// TIA Portal V21 export
// export: Created 2026-08-21T20:18:51.0501839Z, ExportSetting None, DisplayName Totally Integrated Automation Portal, DisplayVersion V21, DisplayName STEP 7 Professional, DisplayVersion V21, DisplayName STEP 7 Safety, DisplayVersion V21, DisplayName Tech WebApplication, DisplayVersion V21, DisplayName WinCC Basic/Comfort/Advanced, DisplayVersion V21, DisplayName WinCC Professional, DisplayVersion V21, DisplayName WinCC Unified, DisplayVersion V21
FUNCTION "V100" : Void   // FC3, FBD
{ S7_Optimized_Access := 'TRUE' }
// stored: SetENOAutomatically false
   VAR_TEMP
      Temp : "DigVal";
      In03 : "DigVal";
      Temp_FF : "DigVal";
      Temp_fromCTRL : "StruCm";
   END_VAR
BEGIN

REGION Network 1: VlvAnL interconnections
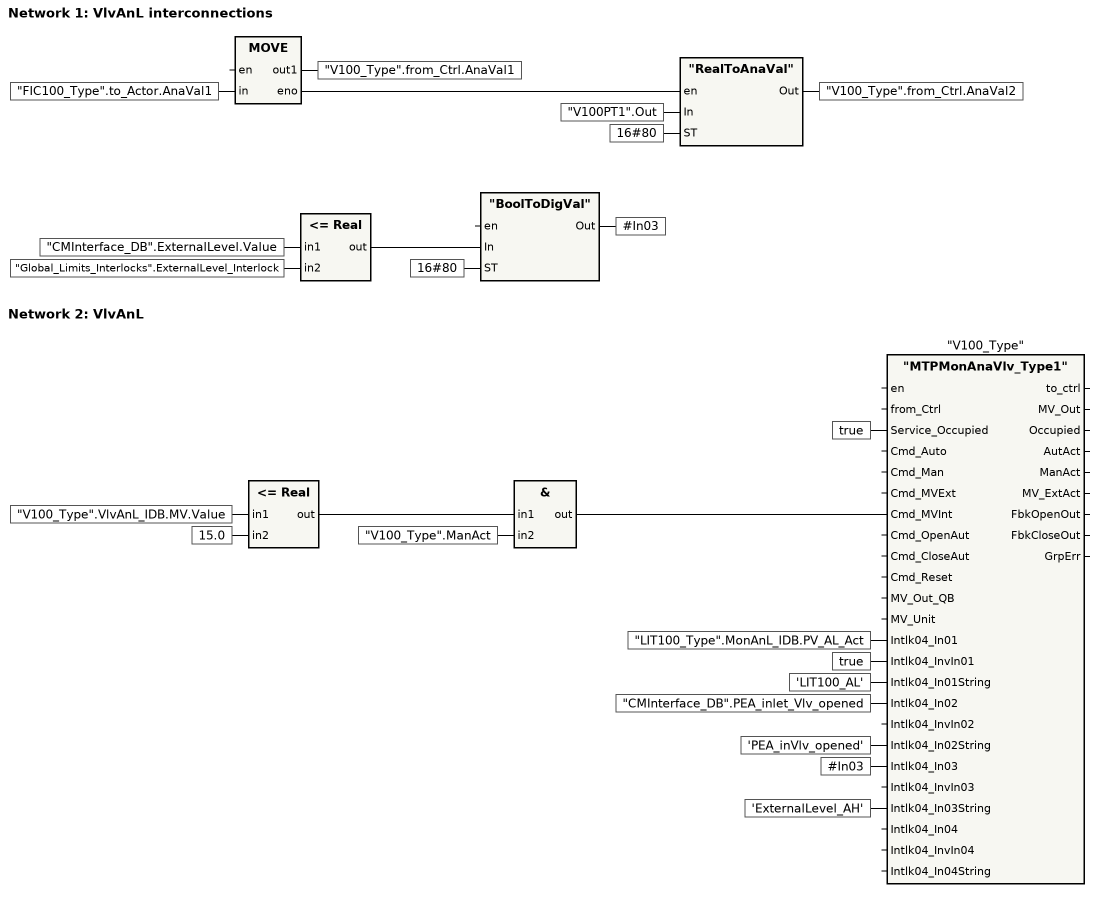
   "V100_Type".from_Ctrl.AnaVal1 := "FIC100_Type".to_Actor.AnaVal1;
   "RealToAnaVal"(In := "V100PT1".Out, ST := 16#80, Out => "V100_Type".from_Ctrl.AnaVal2);
   "BoolToDigVal"(In := "CMInterface_DB".ExternalLevel.Value <= "Global_Limits_Interlocks".ExternalLevel_Interlock,
                  ST := 16#80,
                  Out => #In03);
END_REGION

REGION Network 2: VlvAnL
   "V100_Type"(Service_Occupied := true,   // "MTPMonAnaVlv_Type1"
               Cmd_MVInt := ("V100_Type".VlvAnL_IDB.MV.Value <= 15.0) AND "V100_Type".ManAct,
               Intlk04_In01 := "LIT100_Type".MonAnL_IDB.PV_AL_Act,
               Intlk04_InvIn01 := true,
               Intlk04_In01String := 'LIT100_AL',
               Intlk04_In02 := "CMInterface_DB".PEA_inlet_Vlv_opened,
               Intlk04_In02String := 'PEA_inVlv_opened',
               Intlk04_In03 := #In03,
               Intlk04_In03String := 'ExternalLevel_AH');
END_REGION
END_FUNCTION
